Staubli VAL3: onStart.pgx

public program onStart()
  local num l_nResult
begin
  // call program:loadPROG(0,l_nResult)
  //  if l_nResult!=0
  //    popUpMsg("库加载错误："+toString("",l_nResult))
  //  endIf

  // call refreshproglist()
  call program:getProgList(sProgLsit)
  call refreshlist()

  nPageIndex=0
  nPageNum=roundUp(size(sProgLsit)/49)

  if !isDefined(progTemp:pProgItem[sSelProg])
    sSelProg=""
  endIf
  //
  sPageIndex=toString("",nPageIndex+1)
  sPageNum=toString("",nPageNum)
end
